// TIA Portal V21 export
// export: Created 2026-11-21T13:26:58.7733285Z, ExportSetting WithDefaults, DisplayName Totally Integrated Automation Portal, DisplayVersion V21, DisplayName STEP 7 Professional, DisplayVersion V21, DisplayName STEP 7 Safety, DisplayVersion V21, DisplayName Tech WebApplication, DisplayVersion V21, DisplayName WinCC Basic/Comfort/Advanced, DisplayVersion V21, DisplayName WinCC Unified, DisplayVersion V21
DATA_BLOCK "TankA"   // DB1
VERSION : 0.1
// stored: AutoNumber true, DBAccessibleFromOPCUA true, DBAccessibleFromWebserver true, InstanceOfName Tank, InstanceOfType FB
"Tank"
   // VAR_INPUT
   //    level : Int;
   //    high : Bool;
   //    low : Bool;
   //    state : Int;
   // END_VAR
   // VAR
   //    highAlarm { S7_SetPoint := 'True'} : Program_Alarm;
   //    lowAlarm { S7_SetPoint := 'True'} : Program_Alarm;
   // END_VAR
BEGIN
END_DATA_BLOCK
